(* IEC 61131-3 sources: codesys-to-s7/tests/corpus/C2S7-TYPE-PTR/pos, 1 file *)

(* ---- input.st ---- *)
FUNCTION_BLOCK FB_Case
VAR
    p : POINTER TO INT;
    a : INT;
END_VAR
p := ADR(a);
END_FUNCTION_BLOCK
